// TIA Portal V20 export
// export: Created 2026-10-20T18:54:39.8900098Z, ExportSetting None, DisplayName Totally Integrated Automation Portal, DisplayVersion V20 Update 6, DisplayName TIA Portal Openness, DisplayVersion V20 Update 6, DisplayName TIA Portal Version Control Interface, DisplayVersion V20 Update 6, DisplayName SINAMICS Startdrive Advanced, DisplayVersion V20 SP1, DisplayName SINAMICS Startdrive G130, G150, S120, S150, SINAMICS MV, G220, S200, S210, DisplayVersion V20 SP1, DisplayName SINAMICS Startdrive G110M, G120, G120C, G120D, G120P, G115D, DisplayVersion V20 SP1, DisplayName STEP 7 Professional, DisplayVersion V20 Update 6, DisplayName STEP 7 Safety, DisplayVersion V20 Update 2, DisplayName WinCC Basic/Comfort/Advanced, DisplayVersion V20 Update 6, DisplayName WinCC Unified, DisplayVersion V20 Update 6
VAR_GLOBAL   // PLC tag table "IO_Remote_Panel_1"
   "VTD1 UPPER LIMIT" AT %I118.0 : Bool;
   "VTD1 LOWER LIMIT" AT %I118.3 : Bool;   // TESTED
   "VTD1 PUSH TO ENTER VTD ZONE" AT %I119.4 : Bool;
   "VTD1 PUSH TO EXIT VTD ZONE" AT %I119.5 : Bool;
   "CVTD1 CIRCUIT BREAKER FEEDBACK" AT %I122.0 : Bool;   // TESTED
   "VTD1 CIRCUIT BREAKER FEEDBACK" AT %I122.1 : Bool;   // TESTED
   "CABINET 24V PSU CIRCUIT BREAKER FEEDBACK(1)" AT %I122.2 : Bool;   // IT WILL NEVER GO TO FALSE
   "CABINET COOLING FAN CIRCUIT BREAKER FEEDBACK(1)" AT %I122.3 : Bool;
   "Chain Slack 1 - CH1(1)" AT %I507.0 : Bool;   // TESTED
   "Chain Slack 2 - CH1(1)" AT %I507.1 : Bool;   // TESTED
   "Chain Slack 3 - CH1(1)" AT %I507.2 : Bool;   // TESTED
   "Chain Slack 4 - CH1(1)" AT %I507.3 : Bool;   // TESTED
   "Chain Slack 1 - CH2(1)" AT %I507.4 : Bool;   // TESTED
   "Chain Slack 2 - CH2(1)" AT %I507.5 : Bool;   // TESTED
   "Chain Slack 3 - CH2(1)" AT %I507.6 : Bool;   // TESTED
   "Chain Slack 4 - CH2(1)" AT %I507.7 : Bool;   // TESTED
   "OVERTRAVEL LOWER LIMIT - CH1(1)" AT %I500.0 : Bool;   // TESTED
   "OVERTRAVEL UPPER LIMIT - CH1(1)" AT %I500.1 : Bool;   // Overtravel Upper Limit - CH1
   "E-STOP (CABINET) - CH1(1)" AT %I500.2 : Bool;   // TESTED
   "RESET (CABINET)(1)" AT %I500.3 : Bool;   // TESTED
   "OVERTRAVEL LOWER LIMIT - CH2(1)" AT %I500.4 : Bool;   // Overtravel Lower Limit - CH2
   "OVERTRAVEL UPPER LIMIT - CH2(1)" AT %I500.5 : Bool;   // Overtravel Upper Limit - CH2
   "E-STOP (CABINET) - CH2(1)" AT %I500.6 : Bool;   // E-Stop (Cabinet) - CH2
   "Power Enable Safety Stopper Conveyors (Level 7,8 - Side1) - CH1(1)" AT %Q32.0 : Bool;
   "Power Enable Safety Stopper Conveyors (Level 7,8 - Side1) - CH2(1)" AT %Q32.1 : Bool;
   "Power Enable Safety Stopper Conveyors (Level 7,8 - Side2) - CH1(1)" AT %Q32.2 : Bool;
   "Power Enable Safety Stopper Conveyors (Level 7,8 - Side2) - CH2(1)" AT %Q32.3 : Bool;
   "VTU HOIST BRAKE SAFETY ENABLE 1(1)" AT %Q32.4 : Bool;
   "VTU HOIST BRAKE SAFETY ENABLE 2(1)" AT %Q32.5 : Bool;
   "Power Enable Safety Stopper Conveyors (Level 1,2,3 - Side1) - CH1(1)" AT %Q552.0 : Bool;
   "Power Enable Safety Stopper Conveyors (Level 1,2,3 - Side1) - CH2(1)" AT %Q552.1 : Bool;
   "Power Enable Safety Stopper Conveyors (Level 1,2,3 - Side2) - CH1(1)" AT %Q552.2 : Bool;
   "Power Enable Safety Stopper Conveyors (Level 1,2,3 - Side2) - CH2(1)" AT %Q552.3 : Bool;
   "Power Enable Safety Stopper Conveyors (Level 4,5,6 - Side1) - CH1(1)" AT %Q552.4 : Bool;
   "Power Enable Safety Stopper Conveyors (Level 4,5,6 - Side1) - CH2(1)" AT %Q552.5 : Bool;
   "Power Enable Safety Stopper Conveyors (Level 4,5,6 - Side2) - CH1(1)" AT %Q552.6 : Bool;
   "Power Enable Safety Stopper Conveyors (Level 4,5,6 - Side2) - CH2(1)" AT %Q552.7 : Bool;
   "STO VTD - CH1(1)" AT %Q540.0 : Bool;
   "STO VTD - CH2(1)" AT %Q540.1 : Bool;
   "STO CONVEYOR VTD - CH1(1)" AT %Q540.2 : Bool;
   "STO CONVEYOR VTD - CH2(1)" AT %Q540.3 : Bool;
   "STO CNV VFD (Level 1,2,3 - Side1) - CH1(1)" AT %Q540.4 : Bool;
   "STO CNV VFD (Level 1,2,3 - Side1) - CH2(1)" AT %Q540.5 : Bool;
   "STO CNV VFD (Level 1,2,3 - Side2) - CH1(1)" AT %Q540.6 : Bool;
   "STO CNV VFD (Level 1,2,3 - Side2) - CH2(1)" AT %Q540.7 : Bool;
   "STO CNV VFD (Level 4,5,6 - Side1) - CH1(1)" AT %Q546.0 : Bool;
   "STO CNV VFD (Level 4,5,6 - Side1) - CH2(1)" AT %Q546.1 : Bool;
   "STO CNV VFD (Level 4,5,6 - Side2) - CH1(1)" AT %Q546.2 : Bool;
   "STO CNV VFD (Level 4,5,6 - Side2) - CH2(1)" AT %Q546.3 : Bool;
   "STO CNV VFD (Level 7,8 - Side1) - CH1(1)" AT %Q546.4 : Bool;
   "STO CNV VFD (Level 7,8 - Side1) - CH2(1)" AT %Q546.5 : Bool;
   "STO CNV VFD (Level 7,8 - Side2) - CH1(1)" AT %Q546.6 : Bool;
   "STO CNV VFD (Level 7,8 - Side2) - CH2(1)" AT %Q546.7 : Bool;
   "LIGHT GUARDS C1201 - CH2" AT %I521.4 : Bool;
   "LIGHT GUARDS C1101 - CH1" AT %I521.1 : Bool;
   "LIGHT GUARDS C1101 - CH2" AT %I521.5 : Bool;
   "LIGHT GUARDS C1201 - CH1" AT %I521.0 : Bool;
   "VTD1 SFTY STOPPER CNVS 7,8 - (SIDE 2)" AT %I514.5 : Bool;
   "VTD1 SFTY STOPPER CNVS 7,8 - (SIDE 1)" AT %I514.4 : Bool;
   "SCA 1002 STACK LIGHTS AMBER" AT %Q108.4 : Bool;
   "SCA 1002 STACK LIGHTS GREEN" AT %Q108.5 : Bool;
   "SCA 1002 STACK LIGHTS RED" AT %Q108.6 : Bool;
   "VTD1 SFTY STOPPER CNVS 4,5,6 - (SIDE 2)" AT %I514.3 : Bool;
   "VTD1 SFTY STOPPER CNVS 4,5,6 - (SIDE 1)" AT %I514.2 : Bool;
   "VTD1 DOCKING PINS 2 RETRACT" AT %Q108.1 : Bool;
   "VTD1 DOCKING PINS 1 EXTEND" AT %Q108.2 : Bool;
   "VTD1 SFTY STOPPER CNVS 1,2,3 - (SIDE 1)" AT %I514.0 : Bool;   // SAFETY STOPPER CONVEYORS (1,2,3 - SIDE 1) EDMFEEDBACK
   "VTD1 SFTY STOPPER CNVS 1,2,3 - (SIDE 2)" AT %I514.1 : Bool;
   "VTD1 DOCKING PINS 1 RETRACT" AT %Q108.3 : Bool;
   "EMERGENCY STOP RESET STATUS - ON(1)" AT %Q108.7 : Bool;   // TESTED
   "VTU HOIST BRAKE SAFETY ENABLE EDM FEEDBACK(1)" AT %I514.7 : Bool;
   "C1204_SFTY STOPPER ROTATE" AT %Q101.4 : Bool;
   "C1104_SFTY STOPPER ROTATE" AT %Q105.4 : Bool;
   "C1206_SFTY STOPPER ROTATE" AT %Q102.4 : Bool;
   "C1205_SFTY STOPPER ROTATE" AT %Q102.0 : Bool;
   "C1105_SFTY STOPPER ROTATE" AT %Q106.0 : Bool;
   "C1102_SFTY STOPPER ROTATE" AT %Q104.4 : Bool;
   "C1203_SFTY STOPPER ROTATE" AT %Q101.0 : Bool;
   "C1108_SFTY STOPPER ROTATE" AT %Q107.4 : Bool;
   "C1208_SFTY STOPPER ROTATE" AT %Q103.4 : Bool;
   "C1106_SFTY STOPPER ROTATE" AT %Q106.4 : Bool;
   "C1101_SFTY STOPPER ROTATE" AT %Q104.0 : Bool;
   "C1103_SFTY STOPPER ROTATE" AT %Q105.0 : Bool;   // MOTOR BROKED
   "C1207_SFTY STOPPER ROTATE" AT %Q103.0 : Bool;
   "C1107_SFTY STOPPER ROTATE" AT %Q107.0 : Bool;
   "C1202_SFTY STOPPER ROTATE" AT %Q100.4 : Bool;
   "C1201_SFTY STOPPER ROTATE" AT %Q100.0 : Bool;
   "VTD1 DOCKING PINS 2 EXTEND" AT %Q108.0 : Bool;
   "C1101 CIRCUIT BREAKER FEEDBACK" AT %I121.0 : Bool;   // TESTED
   "C1207 CIRCUIT BREAKER FEEDBACK" AT %I120.6 : Bool;   // TESTED
   "C1108 CIRCUIT BREAKER FEEDBACK" AT %I121.7 : Bool;   // TESTED
   "C1204 CIRCUIT BREAKER FEEDBACK" AT %I120.3 : Bool;   // TESTED
   "C1103 CIRCUIT BREAKER FEEDBACK" AT %I121.2 : Bool;   // TESTED
   "C1206 CIRCUIT BREAKER FEEDBACK" AT %I120.5 : Bool;   // TESTED
   "C1203 CIRCUIT BREAKER FEEDBACK" AT %I120.2 : Bool;   // TESTED
   "C1202 CIRCUIT BREAKER FEEDBACK" AT %I120.1 : Bool;   // TESTED
   "C1205 CIRCUIT BREAKER FEEDBACK" AT %I120.4 : Bool;   // TESTED
   "C1106 CIRCUIT BREAKER FEEDBACK" AT %I121.5 : Bool;   // TESTED
   "C1105 CIRCUIT BREAKER FEEDBACK" AT %I121.4 : Bool;   // TESTED
   "C1201 CIRCUIT BREAKER FEEDBACK" AT %I120.0 : Bool;   // TESTED
   "C1102 CIRCUIT BREAKER FEEDBACK" AT %I121.1 : Bool;   // TESTED
   "C1208 CIRCUIT BREAKER FEEDBACK" AT %I120.7 : Bool;   // TESTED
   "C1107 CIRCUIT BREAKER FEEDBACK" AT %I121.6 : Bool;   // TESTED
   "C1104 CIRCUIT BREAKER FEEDBACK" AT %I121.3 : Bool;   // TESTED
   "GATE_SENSOR_2_CH1(1)" AT %I521.3 : Bool;
   "GATE_SENSOR_1_CH2(1)" AT %I521.6 : Bool;
   "GATE_SENSOR_2_CH2(1)" AT %I521.7 : Bool;
   "GATE_SENSOR_1_CH1(1)" AT %I521.2 : Bool;
END_VAR
